FUNCTION_BLOCK FB_LdCaller
VAR_INPUT
  bEnabled      : BOOL;
  bAuto         : BOOL;
  bManual       : BOOL;
  bJog          : BOOL;
  bFault        : BOOL;
  bPermit       : BOOL;
END_VAR
VAR_OUTPUT
  bRunning      : BOOL;
  bConveyorDone : BOOL;
END_VAR
VAR
  fbConveyor    : FB_Conveyor;
  fbOther       : FB_Sensor;
END_VAR

METHOD MotionCycle
VAR_INPUT
END_VAR
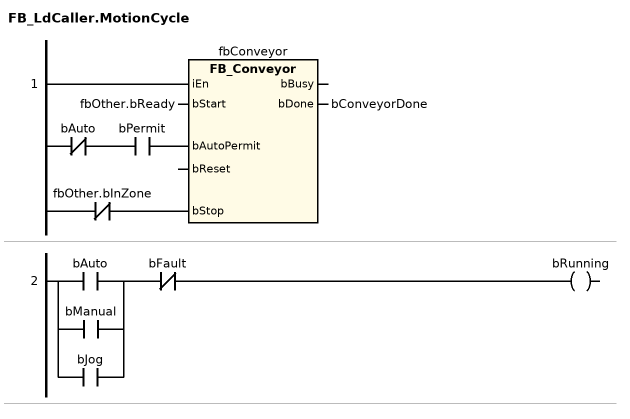
// NETWORK 1
fbConveyor(
    iEn := TRUE,
    bStart := fbOther.bReady,
    bAutoPermit := NOT bAuto AND bPermit,
    bStop := NOT fbOther.bInZone,
    bDone => bConveyorDone); // FB_Conveyor

// NETWORK 2
bRunning := (bAuto OR bManual OR bJog) AND NOT bFault;
END_METHOD

METHOD IdleCycle
VAR_INPUT
END_VAR
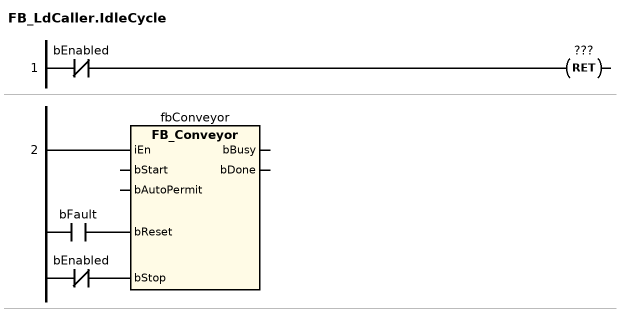
// NETWORK 1
IF NOT bEnabled THEN RETURN; END_IF

// NETWORK 2
fbConveyor(iEn := TRUE, bReset := bFault, bStop := NOT bEnabled); // FB_Conveyor
END_METHOD

END_FUNCTION_BLOCK

(* stored: Version 1.1.0.1, ProductVersion 3.1.4024.12
   POU FB_LdCaller: Id {0a1b2c3d-0000-4000-8000-000000000201}, SpecialFunc None
   Method MotionCycle: Id {0a1b2c3d-0000-4000-8000-000000000202}
   Method IdleCycle: Id {0a1b2c3d-0000-4000-8000-000000000203} *)
